Staubli VAL3: progTemp.pjx

--- progTemp.pjx ---
Parameters version=s8.10.3Cs9_BS2093 stackSize=5000 millimeterUnit=true
Program file=start.pgx
Program file=stop.pgx
Data file=progTemp.dtx
Type name=progItem path=Disk://source/template/progItem/progItem.pjx

--- progTemp.dtx ---
public progItem pProgItem{}
  [Key1]
    progTemplate pProgTemplate
      [0]
        forItem fForItem
          [0]
            bool bIOdisable
            num nLoopValue
            string sForTRAJ
            string sIOindex
        ifItem iIfItem
          [0]
            bool bANDOR[2]
            num nSigIndex[3]
            num nSigType[3]
            num nValue[3]
        num nType
        switchItem sSwitchItem
          [0]
            bool bIOdisable
            num nSwitchValue
            string sIOValue
        string sTRAJname

--- start.pgx ---
program start()
begin
end

--- stop.pgx ---
program stop()
begin
end
